{region 'Documentation'}
(*!
<summary>Checks equality with the expected UDINT value.</summary>
*)
{endregion}
FUNCTION_BLOCK AssertEqual_UDInt EXTENDS AssertionBase
VAR_INPUT
    IN : UDINT; //! Actual value checked or observed by this Assertion.
    Expected : UDINT; //! Reference value for comparison with IN.
END_VAR

SUPER^();

{region 'Documentation'}
(*!
<summary>Check equality with the expected UDINT value.</summary>
*)
{endregion}
METHOD PROTECTED Assert
VAR
    Message : STRING(GVL_Constants.MessageLength);
    ExpectedText : STRING(GVL_Constants.AssertionValueLength);
    ActualText : STRING(GVL_Constants.AssertionValueLength);
END_VAR
IF NOT EvaluationActive THEN
    RETURN;
END_IF;

IF Result = E_Result.Error THEN
    RETURN;
END_IF;

IF Result = E_Result.Failed THEN
    RETURN;
END_IF;

IF IN <> Expected THEN
    ExpectedText := UDINT_TO_STRING(Expected);
    ActualText := UDINT_TO_STRING(IN);
    Message := CONCAT('Assertion failed: values are not equal. Expected = ',
        ExpectedText);
    Message := CONCAT(Message, ', Actual = ');
    Message := CONCAT(Message, ActualText);
    Message := CONCAT(Message, '.');
    Fail(Message := Message);
    RETURN;
END_IF;

Pass();
END_METHOD

END_FUNCTION_BLOCK

(* stored: Version 1.1.0.1
   POU AssertEqual_UDInt: Id {df05908c-bfde-47e0-9412-dd9d9f447ab9}, SpecialFunc None
   Folder Internal: Id {670adf1e-2db4-4765-be6b-db79e5a617b6}
   Method Assert: Id {07b6bbfd-cf8a-4df9-8b77-c2fa21955053} *)
